FUNCTION_BLOCK OUTPUT_PACK (* Migrated from IEC 61131-3 ST *)
  (* Standard: 61499-2 *)
  (* Version 1.0, 2026-11-06, st2fb *)
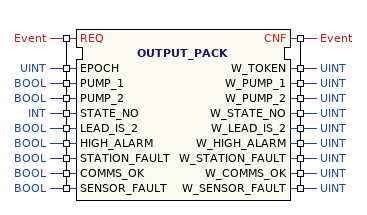
  EVENT_INPUT
    REQ WITH EPOCH, PUMP_1, PUMP_2, STATE_NO, LEAD_IS_2, HIGH_ALARM, STATION_FAULT, COMMS_OK, SENSOR_FAULT;
  END_EVENT
  EVENT_OUTPUT
    CNF WITH W_TOKEN, W_PUMP_1, W_PUMP_2, W_STATE_NO, W_LEAD_IS_2, W_HIGH_ALARM, W_STATION_FAULT, W_COMMS_OK, W_SENSOR_FAULT;
  END_EVENT
  VAR_INPUT
    EPOCH : UINT;
    PUMP_1 : BOOL;
    PUMP_2 : BOOL;
    STATE_NO : INT;
    LEAD_IS_2 : BOOL;
    HIGH_ALARM : BOOL;
    STATION_FAULT : BOOL;
    COMMS_OK : BOOL;
    SENSOR_FAULT : BOOL;
  END_VAR
  VAR_OUTPUT
    W_TOKEN : UINT;
    W_PUMP_1 : UINT;
    W_PUMP_2 : UINT;
    W_STATE_NO : UINT;
    W_LEAD_IS_2 : UINT;
    W_HIGH_ALARM : UINT;
    W_STATION_FAULT : UINT;
    W_COMMS_OK : UINT;
    W_SENSOR_FAULT : UINT;
  END_VAR
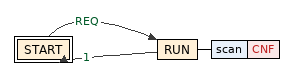
  EC_STATES
    START;
    RUN : scan -> CNF;
  END_STATES
  EC_TRANSITIONS
    START TO RUN := REQ;
    RUN TO START := 1;
  END_TRANSITIONS
  ALGORITHM scan IN ST:
W_TOKEN := EPOCH;
W_PUMP_1 := BOOL_TO_UINT(PUMP_1);
W_PUMP_2 := BOOL_TO_UINT(PUMP_2);
W_STATE_NO := INT_TO_UINT(STATE_NO);
W_LEAD_IS_2 := BOOL_TO_UINT(LEAD_IS_2);
W_HIGH_ALARM := BOOL_TO_UINT(HIGH_ALARM);
W_STATION_FAULT := BOOL_TO_UINT(STATION_FAULT);
W_COMMS_OK := BOOL_TO_UINT(COMMS_OK);
W_SENSOR_FAULT := BOOL_TO_UINT(SENSOR_FAULT);
  END_ALGORITHM
END_FUNCTION_BLOCK
